// TIA Portal V21 export
// export: Created 2026-11-10T07:26:49.4464979Z, ExportSetting WithDefaults, DisplayName Totally Integrated Automation Portal, DisplayVersion V21 Update 3, DisplayName STEP 7 Professional, DisplayVersion V21 Update 3, DisplayName STEP 7 Safety, DisplayVersion V21, DisplayName Tech WebApplication, DisplayVersion V21, DisplayName WinCC Basic/Comfort/Advanced, DisplayVersion V21 Update 3, DisplayName WinCC Unified, DisplayVersion V21 Update 3
FUNCTION_BLOCK "FB_FbdOperands"   // FB6, FBD
{ S7_Optimized_Access := 'TRUE' }
VERSION : 0.1
// stored: AutoNumber true, IsIECCheckEnabled false, IsRetainMemResEnabled false, MemoryReserve 100, SetENOAutomatically false, UDAEnableTagReadback false
   VAR_INPUT
      "a" : Bool;
      ia : Int;
      wa : Word;
   END_VAR
   VAR_OUTPUT
      q : Bool;
      io : Int;
      dout : DInt;
      rout : Real;
      tout : Time;
      sout : String;
   END_VAR
   VAR_IN_OUT
      arr : Array[0..9] of Int;
   END_VAR
   VAR CONSTANT
      cInt : Int := 7;
   END_VAR
BEGIN

REGION Network 1: Absolute address word
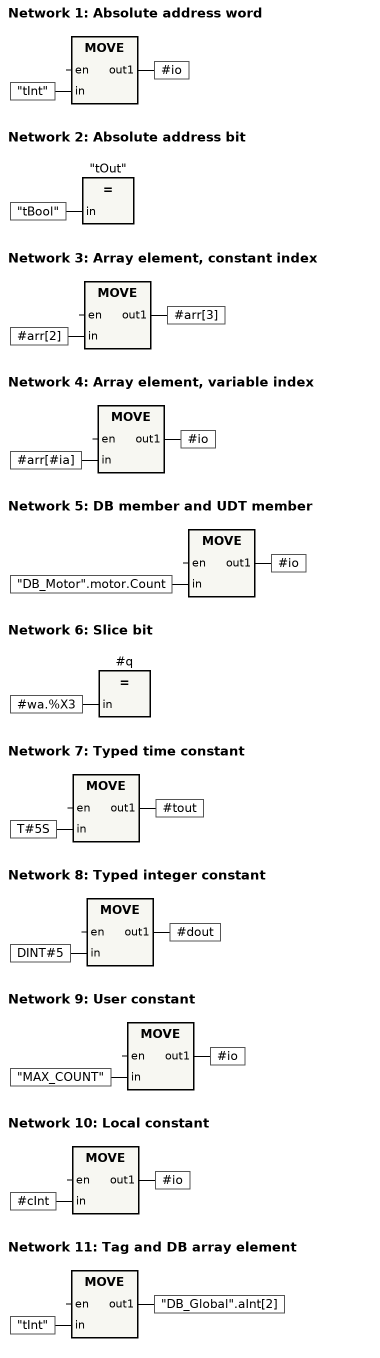
   #io := "tInt";
END_REGION

REGION Network 2: Absolute address bit
   "tOut" := "tBool";
END_REGION

REGION Network 3: Array element, constant index
   #arr[3] := #arr[2];
END_REGION

REGION Network 4: Array element, variable index
   #io := #arr[#ia];
END_REGION

REGION Network 5: DB member and UDT member
   #io := "DB_Motor".motor.Count;
END_REGION

REGION Network 6: Slice bit
   #q := #wa.%X3;
END_REGION

REGION Network 7: Typed time constant
   #tout := T#5S;
END_REGION

REGION Network 8: Typed integer constant
   #dout := DINT#5;
END_REGION

REGION Network 9: User constant
   #io := "MAX_COUNT";
END_REGION

REGION Network 10: Local constant
   #io := #cInt;
END_REGION

REGION Network 11: Tag and DB array element
   "DB_Global".aInt[2] := "tInt";
END_REGION

REGION Network 12: Real literal
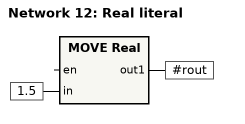
   #rout := 1.5;
END_REGION
END_FUNCTION_BLOCK
